INTERFACE I_CustomStationInterface

PROPERTY pressedAbortButton  : BOOL
GET
END_GET
END_PROPERTY

END_INTERFACE

(* stored: Version 1.1.0.1, ProductVersion 3.1.4024.12
   Itf I_CustomStationInterface: Id {9135faed-838e-4c82-9a7a-8ea69bc3c123}
   Property pressedAbortButton: Id {067a4613-d0b4-408d-a0cf-5f6fe8eca99d}
   Get Get: Id {8240dc48-d178-42ab-b318-b1f727331493} *)
